// Mock of the focus axis (I_Focus) for the telescope state machine tests: enabled = ready and calibrated at once (the telescope never sets HomeAxis), the
// position follows the target at once. Status only, no motion model.
FUNCTION_BLOCK FB_FocusMock IMPLEMENTS BROTLib.I_Focus
VAR
	bEn		: BOOL;
	bCal	: BOOL;
	bHome	: BOOL;
	bNeg	: BOOL;
	bPos	: BOOL;
	fPos	: LREAL;
	fTarget	: LREAL;
	fVel	: LREAL;
	nStop	: INT;		// number of Stop() calls
END_VAR

IF bEn THEN
	bCal := TRUE;
END_IF
fPos := fTarget;

METHOD Stop : BOOL
nStop := nStop + 1;
Stop := TRUE;
END_METHOD

PROPERTY MinPosition : LREAL
GET
MinPosition := -1.0E6;
END_GET
END_PROPERTY

PROPERTY MaxPosition : LREAL
GET
MaxPosition := 1.0E6;
END_GET
END_PROPERTY

METHOD Reset : BOOL
Reset := TRUE;
END_METHOD

PROPERTY ActualPosition : LREAL
GET
ActualPosition := fPos;
END_GET
SET
fPos := ActualPosition;
END_SET
END_PROPERTY

PROPERTY Busy : BOOL
GET
Busy := FALSE;
END_GET
END_PROPERTY

PROPERTY Calibrated : BOOL
GET
Calibrated := bCal;
END_GET
END_PROPERTY

PROPERTY Enable : BOOL
GET
Enable := bEn;
END_GET
SET
bEn := Enable;
END_SET
END_PROPERTY

PROPERTY Error : BOOL
GET
Error := FALSE;
END_GET
END_PROPERTY

PROPERTY ErrorID : UDINT
GET
ErrorID := 0;
END_GET
END_PROPERTY

PROPERTY HomeAxis : BOOL
GET
HomeAxis := bHome;
END_GET
SET
bHome := HomeAxis;
END_SET
END_PROPERTY

PROPERTY InNegLimit : BOOL
GET
InNegLimit := FALSE;
END_GET
END_PROPERTY

PROPERTY InPosLimit : BOOL
GET
InPosLimit := FALSE;
END_GET
END_PROPERTY

PROPERTY MoveNeg : BOOL
GET
MoveNeg := bNeg;
END_GET
SET
bNeg := MoveNeg;
END_SET
END_PROPERTY

PROPERTY MovePos : BOOL
GET
MovePos := bPos;
END_GET
SET
bPos := MovePos;
END_SET
END_PROPERTY

PROPERTY Position : LREAL
GET
Position := fTarget;
END_GET
SET
fTarget := Position;
END_SET
END_PROPERTY

PROPERTY Ready : BOOL
GET
Ready := bEn;
END_GET
END_PROPERTY

PROPERTY Velocity : LREAL
GET
Velocity := fVel;
END_GET
SET
fVel := Velocity;
END_SET
END_PROPERTY

END_FUNCTION_BLOCK

(* stored: Version 1.1.0.1, ProductVersion 3.1.4024.15
   POU FB_FocusMock: Id {5fdf5a9a-cc47-484b-b66c-dbdc86e8cac2}, SpecialFunc None
   Method Stop: Id {23bdd15b-5914-43f8-a4ab-1ddba78da4a7}
   Property MinPosition: Id {5d6ac3d9-931e-465f-85f9-3defb9d0eb84}
   Get Get: Id {088902ba-9239-4fb9-8d7a-53d6f6cd726c}
   Property MaxPosition: Id {278fefd5-d20e-4b37-8369-b61d776d023f}
   Get Get: Id {dcffa58f-8457-49a9-a82b-e5d4f2db68f5}
   Method Reset: Id {14e9fc07-28bd-416d-89a8-915cece929c7}
   Property ActualPosition: Id {1a1423fd-de3c-46bb-9a00-026fe8bbcf63}
   Get Get: Id {e8baa86d-f60c-40f4-a253-ac333fc9acfb}
   Set Set: Id {f516f653-7e75-44fd-a6ef-1ecb90d940d1}
   Property Busy: Id {fac01a2e-5806-47d6-8e56-d26f2542c24a}
   Get Get: Id {85dd49f5-6cbd-4e15-baff-c3f0242c8549}
   Property Calibrated: Id {063c579e-92d0-4642-ba8b-29b00f044579}
   Get Get: Id {463cd35a-c468-42d7-bddb-8728ecca8523}
   Property Enable: Id {f5761f92-7d0d-4820-99f2-cccd25a13541}
   Get Get: Id {cd71e71b-1565-40f7-b7f3-35a6f2719038}
   Set Set: Id {edc46e04-4bfa-4e20-9123-3cf4493fa673}
   Property Error: Id {e6a5b0eb-7e80-470b-b7ce-5bbac5d77f2b}
   Get Get: Id {a05e5e81-bdfd-469d-8192-c521ca62a37d}
   Property ErrorID: Id {4592d737-db73-4bd4-bbc7-77f6ecbd80c5}
   Get Get: Id {df82a7dd-d67c-47cb-bde4-5b2d4b9bce4d}
   Property HomeAxis: Id {81f497f9-3ab3-440d-9c19-f555c1ac29b5}
   Get Get: Id {17c9df60-8f06-466d-9b1c-6f0fc5ea1529}
   Set Set: Id {45b1fdad-7075-481b-a3c1-b31da2264621}
   Property InNegLimit: Id {9a20bb8e-5943-43a3-9ecc-570004978da3}
   Get Get: Id {6c666f07-6f98-491c-9784-448cff620f7e}
   Property InPosLimit: Id {2af08350-a65f-44a1-b036-d3622cdf45de}
   Get Get: Id {e03f0a88-6a3a-43bc-80cc-517b6d9471e3}
   Property MoveNeg: Id {3f1e0455-2e10-4f97-b91e-3839debaa5c0}
   Get Get: Id {e9ef14b5-a4c0-4454-855f-25bfc4edeee4}
   Set Set: Id {ff8707b6-531b-4550-9841-d5e91393b0d4}
   Property MovePos: Id {4e5a3388-e926-4c60-9021-1bacdef16e67}
   Get Get: Id {df4e8889-26e0-46aa-8099-8aa25760fab9}
   Set Set: Id {22d332c7-8c4a-4bda-8e67-6a78d82f310a}
   Property Position: Id {3997f07a-6f54-4add-8f61-68eebf5349c4}
   Get Get: Id {90545b29-a4ed-45ce-80cb-a8e6bbd5d1a5}
   Set Set: Id {d2f183f8-ce0a-4b29-ab26-b85b6dfdc1ac}
   Property Ready: Id {8dd3f665-be74-4b4a-8b31-59a0c7864d76}
   Get Get: Id {28c6dc8d-7667-4ce0-bbda-dc4392d544b8}
   Property Velocity: Id {f0d5095e-c392-423e-865e-ecad1c412313}
   Get Get: Id {bde2de11-7389-4b00-b868-4421f5d46e99}
   Set Set: Id {92003e7d-811e-490b-a911-167ccac59e86} *)
